(*
SPDX-FileCopyrightText: c 2026 Oleksandr Tiutyk <trofimich@gmail.com>
SPDX-License-Identifier: MIT
License: https://opensource.org/license/mit
*)

(*!
<summary>Groups byte-list operations with dynamically allocated storage.</summary>
<description>
Owns the independent child instances and their fixed registration array. Use from one PLC task at a stable address.
</description>
*)

{attribute 'no_assign'}
{attribute 'no_explicit_call' := 'do not call this function block directly'}
FUNCTION_BLOCK DynamicByteListTestGroup EXTENDS TOF_Testing.TestGroup<6>
VAR_STAT
	{attribute 'hide'}
	_ClassName : STRING := __POUNAME();
END_VAR
VAR
	_LoadFromAny : ByteListLoadFromAnyTest(name := "LoadFromAny", parent := THIS^, useDynamicStorage := TRUE);
	_GetAndSet : ByteListIndexedAccessTest(name := "GetAndSet", parent := THIS^, useDynamicStorage := TRUE);
	_Find : ByteListFindTest(name := "Find", parent := THIS^, useDynamicStorage := TRUE);
	_Remove : ByteListRemoveValueTest(name := "Remove", parent := THIS^, useDynamicStorage := TRUE);
	_RemoveAt : ByteListRemoveRangeTest(name := "RemoveAt", parent := THIS^, useDynamicStorage := TRUE);
	_Clear : ByteListClearTest(name := "Clear", parent := THIS^, useDynamicStorage := TRUE);

	_Children : ARRAY [0.._ChildCount - 1] OF TOF_Testing.ITestElement :=
	[
		_LoadFromAny,
		_GetAndSet,
		_Find,
		_Remove,
		_RemoveAt,
		_Clear
	];
END_VAR

//! <summary>Borrows the fixed child array. Callers must not modify it.</summary>
{attribute 'monitoring' := 'call'}
PROPERTY Children : REFERENCE TO ARRAY [0.._ChildCount - 1] OF TOF_Testing.ITestElement
GET
Children REF= _Children;
END_GET
END_PROPERTY

//! <summary>Borrows the concrete class name. Callers must not modify it.</summary>
{attribute 'monitoring' := 'call'}
PROPERTY ClassName : REFERENCE TO STRING
GET
ClassName REF= _ClassName;
END_GET
END_PROPERTY

//! <summary>Borrows the compiler-initialized namespace name. Callers must not modify it.</summary>
{attribute 'monitoring' := 'call'}
PROPERTY NamespaceName : REFERENCE TO STRING
GET
NamespaceName REF= CurrentNamespace.Name;
END_GET
END_PROPERTY

//! <summary>Reports the concrete instance size in bytes.</summary>
{attribute 'monitoring' := 'call'}
PROPERTY SelfSize : ULINT
GET
SelfSize := XSIZEOF(THIS^);
END_GET
END_PROPERTY

END_FUNCTION_BLOCK

(* stored: Version 1.1.0.1
   POU DynamicByteListTestGroup: Id {e04ef593-b7dd-4488-9412-785966fa705a}, SpecialFunc None
   Property Children: Id {df27839e-4f32-4539-8f00-f5c5461f5a15}
   Get Get: Id {d2ec162c-c2c5-4191-8167-107fe406f129}
   Property ClassName: Id {3c181f2d-038f-4b79-9680-ada7b1a37c18}
   Get Get: Id {debc8bae-ff16-4f4d-8657-42c27c3d1eca}
   Property NamespaceName: Id {c1411af5-c5a2-4549-a59a-f929ecbe09cd}
   Get Get: Id {e28d5fb1-366c-416d-ab46-9be333361efd}
   Property SelfSize: Id {a54ab3b9-22c9-45d8-ba3b-ebf5ab131295}
   Get Get: Id {6448cdf5-0c1e-49e6-ad67-246f9aa7809c} *)
